(* IEC 61131-3 sources: plcassist-cli/packages/volt-lsp-iec/test-corpus/awa-palletizer/Device/Plc Logic/Application/Library Manager/VisuDialogs, 50 files *)

(* ---- DIALOG_CONSTANTS.gvl ---- *)
VAR_GLOBAL
	USERNAME_LABEL_DEFAULT : STRING := 'User';
	PASSWORD_LABEL_DEFAULT : STRING := 'Password';
	LOGIN_DIALOG_NAME : STRING := 'VisuDialogs.Login';
	PASSWORD_CHAR : STRING(1) := '*';
	CHAR_ASTERISK : BYTE := 42;
	CHAR_POINT : BYTE := 46;
	CHAR_SLASH : BYTE := 47;
	CHAR_BACKSLASH : BYTE := 92;
	ERR_DIR_NOT_FOUND : DWORD := 4000;
	ITFID_IGENERALCOMMAND : DWORD := 2;
	VISUDIALOGS_VERSION_ATLEAST_3_5_5 : INT := 0;
END_VAR

(* ---- DIALOG_VARIABLES.gvl ---- *)
VAR_GLOBAL
	G_FILELISTPROVIDER : Visu_FbFileListProvider;
	G_VISUDIALOGSCOMMANDS : Visu_DialogCommands;
END_VAR

(* ---- DIALOG_VARIABLES_EXP.gvl ---- *)
VAR_GLOBAL
	G_XEXP : BOOL;
END_VAR

(* ---- GVL_SORTEDFILELIST.gvl ---- *)
VAR_GLOBAL
	FILEELEMENTFACTORY : SortedDirectoryFileElementFactory;
	SORTEDLISTFACTORY : COL.SortedListFactory;
END_VAR

(* ---- IDIRECTORYFILEELEMENT.itf ---- *)
INTERFACE IDIRECTORYFILEELEMENT
END_INTERFACE

(* ---- IFILELISTPROVIDER.itf ---- *)
INTERFACE IFILELISTPROVIDER
END_INTERFACE

METHOD INITIALIZE : BOOL
VAR_INPUT
	STDIRECTORY : STRING(255);
	STFILTER : STRING;
	STFILEIN : STRING;
	STTITLE : STRING;
	IROWCOUNT : INT;
	BBROWSEDIRECTORY : BOOL;
	BTOUCH : BOOL;
END_VAR
END_METHOD

METHOD NEXT : BOOL
END_METHOD

METHOD PREVIOUS : BOOL
END_METHOD

(* ---- DIALOGCHECKINIT.fun ---- *)
FUNCTION DIALOGCHECKINIT : BOOL
VAR_IN_OUT
	STVALUE : STRING;
	STOUTPUT : STRING;
	BINIT : BOOL;
END_VAR
END_FUNCTION

(* ---- DIALOGCHECKINITFOREXPONENTIAL.fun ---- *)
FUNCTION DIALOGCHECKINITFOREXPONENTIAL : BOOL
VAR_INPUT
	STVALUE : STRING;
END_VAR
VAR_IN_OUT
	BINIT : BOOL;
END_VAR
END_FUNCTION

(* ---- DIALOGCHECKINITFOREXPONENTIALW.fun ---- *)
FUNCTION DIALOGCHECKINITFOREXPONENTIALW : BOOL
VAR_INPUT
	WSTVALUE : WSTRING;
END_VAR
VAR_IN_OUT
	BINIT : BOOL;
END_VAR
END_FUNCTION

(* ---- DIALOGCHECKINITW.fun ---- *)
FUNCTION DIALOGCHECKINITW : BOOL
VAR_IN_OUT
	WSTVALUE : WSTRING;
	WSTOUTPUT : WSTRING;
	BINIT : BOOL;
END_VAR
END_FUNCTION

(* ---- VISUDLG_CHECKEDAPPEND.fun ---- *)
FUNCTION VISUDLG_CHECKEDAPPEND : BOOL
VAR_INPUT
	BPASSWORD : BOOL;
	CTOAPPEND : STRING(1);
END_VAR
VAR_IN_OUT
	STOUTPUTVALUE : STRING;
	STVARIABLEVALUE : STRING;
	BINIT : BOOL;
END_VAR
END_FUNCTION

(* ---- VISUDLG_CHECKEDAPPENDEXP.fun ---- *)
FUNCTION VISUDLG_CHECKEDAPPENDEXP : BOOL
VAR_INPUT
	BPASSWORD : BOOL;
END_VAR
VAR_IN_OUT
	STOUTPUTVALUE : STRING;
	STVARIABLEVALUE : STRING;
	BINIT : BOOL;
END_VAR
END_FUNCTION

(* ---- VISUDLG_CHECKEDAPPENDW.fun ---- *)
FUNCTION VISUDLG_CHECKEDAPPENDW : BOOL
VAR_INPUT
	BPASSWORD : BOOL;
	CTOAPPEND : WSTRING(1);
END_VAR
VAR_IN_OUT
	WSTOUTPUTVALUE : WSTRING;
	WSTVARIABLEVALUE : WSTRING;
	BINIT : BOOL;
END_VAR
END_FUNCTION

(* ---- VISUDLG_CHECKEDBACK.fun ---- *)
FUNCTION VISUDLG_CHECKEDBACK : BOOL
VAR_IN_OUT
	STOUTPUTVALUE : STRING;
	STVARIABLEVALUE : STRING;
	BINIT : BOOL;
END_VAR
END_FUNCTION

(* ---- VISUDLG_CHECKEDBACKW.fun ---- *)
FUNCTION VISUDLG_CHECKEDBACKW : BOOL
VAR_IN_OUT
	WSTOUTPUTVALUE : WSTRING;
	WSTVARIABLEVALUE : WSTRING;
	BINIT : BOOL;
END_VAR
END_FUNCTION

(* ---- VISUDLG_CHECKEDCHANGENUMBERFORMAT.fun ---- *)
FUNCTION VISUDLG_CHECKEDCHANGENUMBERFORMAT : BOOL
VAR_INPUT
	BPASSWORD : BOOL;
	STCLICKEDRADIO : STRING;
END_VAR
VAR_IN_OUT
	STOUTPUTVALUE : STRING;
	STVARIABLEVALUE : STRING;
	STMIN : STRING;
	STMAX : STRING;
	IFORMATVALUE : INT;
END_VAR
END_FUNCTION

(* ---- VISUDLG_CHECKEDCHANGESIGN.fun ---- *)
FUNCTION VISUDLG_CHECKEDCHANGESIGN : BOOL
VAR_INPUT
	BPASSWORD : BOOL;
END_VAR
VAR_IN_OUT
	STOUTPUTVALUE : STRING;
	STVARIABLEVALUE : STRING;
	BINIT : BOOL;
END_VAR
END_FUNCTION

(* ---- VISUDLG_CHECKEDCHANGESIGNEXTENDED.fun ---- *)
FUNCTION VISUDLG_CHECKEDCHANGESIGNEXTENDED : BOOL
VAR_INPUT
	BPASSWORD : BOOL;
	IFORMATVALUE : INT;
END_VAR
VAR_IN_OUT
	STOUTPUTVALUE : STRING;
	STVARIABLEVALUE : STRING;
	BINIT : BOOL;
END_VAR
END_FUNCTION

(* ---- VISUDLG_CHECKEDCLEAR.fun ---- *)
FUNCTION VISUDLG_CHECKEDCLEAR : BOOL
VAR_IN_OUT
	STOUTPUTVALUE : STRING;
	STVARIABLEVALUE : STRING;
	FLAGS : DWORD;
END_VAR
END_FUNCTION

(* ---- VISUDLG_CHECKEDEXPFLOATFORMATSWITCH.fun ---- *)
FUNCTION VISUDLG_CHECKEDEXPFLOATFORMATSWITCH : BOOL
VAR_INPUT
	BPASSWORD : BOOL;
END_VAR
VAR_IN_OUT
	STOUTPUTVALUE : STRING;
	STVARIABLEVALUE : STRING;
END_VAR
END_FUNCTION

(* ---- VISUDLG_GETPASSWORDSTRING.fun ---- *)
FUNCTION VISUDLG_GETPASSWORDSTRING : STRING
VAR_INPUT
	STORG : STRING;
END_VAR
END_FUNCTION

(* ---- VISUDLG_PROCESSCHANGENUMBERFORMAT.fun ---- *)
FUNCTION VISUDLG_PROCESSCHANGENUMBERFORMAT : BOOL
VAR_INPUT
	BPASSWORD : BOOL;
	STCLICKEDRADIO : STRING;
END_VAR
VAR_IN_OUT
	STOUTPUTVALUE : STRING;
	STVARIABLEVALUE : STRING;
	STMIN : STRING;
	STMAX : STRING;
	IFORMATVALUE : INT;
	ICARETPOSITION : INT;
	ISELECTIONSTART : INT;
	ISELECTIONEND : INT;
END_VAR
END_FUNCTION

(* ---- VISUDLG_PROCESSCHANGESIGN.fun ---- *)
FUNCTION VISUDLG_PROCESSCHANGESIGN : BOOL
VAR_INPUT
	BPASSWORD : BOOL;
END_VAR
VAR_IN_OUT
	STOUTPUTVALUE : STRING;
	STVARIABLEVALUE : STRING;
	ICARETPOSITION : INT;
	ISELECTIONSTART : INT;
	ISELECTIONEND : INT;
END_VAR
END_FUNCTION

(* ---- VISUDLG_PROCESSCHANGESIGNEXTENDED.fun ---- *)
FUNCTION VISUDLG_PROCESSCHANGESIGNEXTENDED : BOOL
VAR_INPUT
	BPASSWORD : BOOL;
	IFORMATVALUE : INT;
END_VAR
VAR_IN_OUT
	STOUTPUTVALUE : STRING;
	STVARIABLEVALUE : STRING;
	ICARETPOSITION : INT;
	ISELECTIONSTART : INT;
	ISELECTIONEND : INT;
	BINIT : BOOL;
END_VAR
END_FUNCTION

(* ---- VISUDLG_PROCESSCLEAR.fun ---- *)
FUNCTION VISUDLG_PROCESSCLEAR : BOOL
VAR_IN_OUT
	STOUTPUTVALUE : STRING;
	STVARIABLEVALUE : STRING;
	FLAGS : DWORD;
	ICARETPOSITION : INT;
	ISELECTIONSTART : INT;
	ISELECTIONEND : INT;
END_VAR
END_FUNCTION

(* ---- VISUDLG_PROCESSEXP.fun ---- *)
FUNCTION VISUDLG_PROCESSEXP : BOOL
VAR_INPUT
	BPASSWORD : BOOL;
END_VAR
VAR_IN_OUT
	STOUTPUTVALUE : STRING;
	STVARIABLEVALUE : STRING;
	ICARETPOSITION : INT;
	ISELECTIONSTART : INT;
	ISELECTIONEND : INT;
	BINIT : BOOL;
END_VAR
END_FUNCTION

(* ---- VISUDLG_PROCESSEXPFLOATFORMATSWITCH.fun ---- *)
FUNCTION VISUDLG_PROCESSEXPFLOATFORMATSWITCH : BOOL
VAR_INPUT
	BPASSWORD : BOOL;
END_VAR
VAR_IN_OUT
	STOUTPUTVALUE : STRING;
	STVARIABLEVALUE : STRING;
	ICARETPOSITION : INT;
	ISELECTIONSTART : INT;
	ISELECTIONEND : INT;
	BINIT : BOOL;
END_VAR
END_FUNCTION

(* ---- VISUDLG_SETERRORCOLOR.fun ---- *)
FUNCTION VISUDLG_SETERRORCOLOR : DWORD
VAR_INPUT
	BERROR : BOOL;
END_VAR
END_FUNCTION

(* ---- VISUDLG_UTF8PASSWORDCARETPOSITION.fun ---- *)
FUNCTION VISUDLG_UTF8PASSWORDCARETPOSITION : INT
VAR_INPUT
	IRUNELEN : INT;
	STVARIABLE : STRING;
END_VAR
END_FUNCTION

(* ---- VISUDLG_UTF8RUNELEN.fun ---- *)
FUNCTION VISUDLG_UTF8RUNELEN : INT
VAR_INPUT
	STVARIABLEVALUE : STRING;
	IINDEX : INT;
END_VAR
END_FUNCTION

(* ---- VISUDLGUTIL_CLOSENUMPADEXTENDED.fun ---- *)
FUNCTION VISUDLGUTIL_CLOSENUMPADEXTENDED : BOOL
VAR_INPUT
	FLAGS : DWORD;
END_VAR
VAR_IN_OUT
	STOUTPUTVALUE : STRING;
	STVARIABLEVALUE : STRING;
	STMIN : STRING;
	STMAX : STRING;
	IFORMATVALUE : INT;
	BINITFORMATVALUE : BOOL;
END_VAR
END_FUNCTION

(* ---- VISUDLGUTIL_CLOSENUMPADEXTENDED2.fun ---- *)
FUNCTION VISUDLGUTIL_CLOSENUMPADEXTENDED2 : BOOL
VAR_INPUT
	FLAGS : DWORD;
END_VAR
VAR_IN_OUT
	STOUTPUTVALUE : STRING;
	STVARIABLEVALUE : STRING;
	STMIN : STRING;
	STMAX : STRING;
	IFORMATVALUE : INT;
	BINITFORMATVALUE : BOOL;
	ICARETPOSITION : INT;
	ISELECTIONSTART : INT;
	ISELECTIONEND : INT;
END_VAR
END_FUNCTION

(* ---- VISUDLGUTIL_FORMATEXPTOG.fun ---- *)
FUNCTION VISUDLGUTIL_FORMATEXPTOG : STRING
VAR_INPUT
	STVALUE : STRING;
END_VAR
END_FUNCTION

(* ---- VISUDLGUTIL_FORMATVALUETODEC.fun ---- *)
FUNCTION VISUDLGUTIL_FORMATVALUETODEC : STRING
VAR_INPUT
	STVARIABLEVALUE : STRING;
END_VAR
END_FUNCTION

(* ---- VISUDLGUTIL_FORMATVALUETOHEX.fun ---- *)
FUNCTION VISUDLGUTIL_FORMATVALUETOHEX : STRING
VAR_INPUT
	STVARIABLEVALUE : STRING;
END_VAR
END_FUNCTION

(* ---- VISUDLGUTIL_INITVALUEFROMFLAGS.fun ---- *)
FUNCTION VISUDLGUTIL_INITVALUEFROMFLAGS : INT
VAR_INPUT
	FLAGS : DWORD;
END_VAR
VAR_IN_OUT
	BINITFORMATVALUE : BOOL;
	IFORMATVALUE : INT;
END_VAR
END_FUNCTION

(* ---- VISUDLGUTIL_ISDIALOGOPEN.fun ---- *)
FUNCTION VISUDLGUTIL_ISDIALOGOPEN : BOOL
VAR_INPUT
	LOGINDIALOG : VisuElems.VisuElemBase.IVisualisationDialog;
	PVISUCLIENT : POINTER TO VisuElems.VisuElemBase.VisuStructClientData;
	DLGMAN : VisuElems.VisuElemBase.IDialogManager;
END_VAR
END_FUNCTION

(* ---- VISUDLGUTIL_SETBINITFORMATVALUE.fun ---- *)
FUNCTION VISUDLGUTIL_SETBINITFORMATVALUE : BOOL
VAR_INPUT
	STNEWVALUE : STRING;
END_VAR
VAR_IN_OUT
	BINITFORMATVALUE : BOOL;
END_VAR
END_FUNCTION

(* ---- VISUDLGUTIL_UPDATEOUTPUTVALUE.fun ---- *)
FUNCTION VISUDLGUTIL_UPDATEOUTPUTVALUE : BOOL
VAR_INPUT
	BPASSWORD : BOOL;
END_VAR
VAR_IN_OUT
	STOUTPUTVALUE : STRING;
	STVARIABLEVALUE : STRING;
END_VAR
END_FUNCTION

(* ---- GLOBALTEXTLIST.fb ---- *)
FUNCTION_BLOCK GLOBALTEXTLIST
VAR
	M_TEXTLISTFILE : STRING(255);
	_STNAMESPACE : STRING;
END_VAR
END_FUNCTION_BLOCK

(* ---- IMAGEPOOLDIALOGS.fb ---- *)
FUNCTION_BLOCK IMAGEPOOLDIALOGS
VAR
	M_STNAMESPACE : STRING(80);
	M_STHELPVARID : STRING;
	M_STHELPVARPATH : STRING(255);
	M_STHELP : STRING;
	M_REGISTERIMAGES : BOOL := TRUE;
END_VAR
END_FUNCTION_BLOCK

METHOD FB_INIT : BOOL
VAR_INPUT
	BINITRETAINS : BOOL;
	BINCOPYCODE : BOOL;
END_VAR
END_METHOD

METHOD FB_REINIT : BOOL
END_METHOD

METHOD FB_EXIT : BOOL
VAR_INPUT
	BINCOPYCODE : BOOL;
END_VAR
END_METHOD

(* ---- MINMAXLABELS.fb ---- *)
FUNCTION_BLOCK MINMAXLABELS
VAR
	M_TEXTLISTFILE : STRING(255);
	_STNAMESPACE : STRING;
END_VAR
END_FUNCTION_BLOCK

(* ---- SORTEDDIRECTORYFILEELEMENT.fb ---- *)
FUNCTION_BLOCK SORTEDDIRECTORYFILEELEMENT EXTENDS InstanceBase
VAR
	STFILENAME : STRING;
	DIRINFO : DirInfo;
	DIRECTORYINFO : POINTER TO DirInfo;
	FILENAME : POINTER TO STRING;
END_VAR
END_FUNCTION_BLOCK

METHOD DISPOSE : BOOL
END_METHOD

METHOD PRVINSTINIT : FBF.Error
VAR_INPUT
	ITFDATA : FBF.IData;
END_VAR
END_METHOD

METHOD ELEMENTCOMPARETO : INT
VAR_INPUT
	ITFELEMENT : COL.IElement;
END_VAR
END_METHOD

METHOD ELEMENTEQUALS : BOOL
VAR_INPUT
	ITFELEMENT : COL.IElement;
END_VAR
END_METHOD

METHOD ELEMENTHASHCODE : LINT
END_METHOD

(* ---- SORTEDDIRECTORYFILEELEMENTDATA.fb ---- *)
FUNCTION_BLOCK SORTEDDIRECTORYFILEELEMENTDATA EXTENDS InstanceData
VAR_INPUT
	STFILENAME : STRING;
	DIRINFO : DirInfo;
END_VAR
END_FUNCTION_BLOCK

(* ---- SORTEDDIRECTORYFILEELEMENTFACTORY.fb ---- *)
FUNCTION_BLOCK SORTEDDIRECTORYFILEELEMENTFACTORY EXTENDS FactoryBase
VAR
	PRVINSTCOUNT : CAA.COUNT;
	PRVINSTPOOLEXTENDSFACTOR : USINT;
	PRVINSTSIZE : CAA.SIZE;
END_VAR
END_FUNCTION_BLOCK

METHOD CREATE : IDirectoryFileElement
VAR_INPUT
	STFILENAME : STRING;
	DIRINFO : DirInfo;
END_VAR
VAR_OUTPUT
	EERROR : FBF.ERROR;
END_VAR
END_METHOD

(* ---- VISU_DIALOGCOMMANDS.fb ---- *)
FUNCTION_BLOCK VISU_DIALOGCOMMANDS
VAR
	_CMDOPENFILEDIALOG : Visu_FbOpenFileDialog;
END_VAR
END_FUNCTION_BLOCK

METHOD FB_INIT
VAR_INPUT
	BINITRETAINS : BOOL;
	BINCOPYCODE : BOOL;
END_VAR
END_METHOD

METHOD REGISTERCOMMANDS : BOOL
VAR_INPUT
	COMMANDMANAGER : VisuElems.ICommandManager2;
END_VAR
END_METHOD

(* ---- VISU_FBDIALOGLOGINPROVIDER.fb ---- *)
FUNCTION_BLOCK VISU_FBDIALOGLOGINPROVIDER
VAR
	_STPASSWORD : STRING;
	_STUSERNAME : STRING;
	_CREDENTIALS : Visu_UserPasswordCredentials;
	_STTITLEPREFIX : STRING;
	_STCURRENTDATASOURCE : STRING;
	_STUSERLABELTEXT : STRING;
	_STPASSWORDLABELTEXT : STRING;
	_UXIPROVIDINGCREDENTIALSFOR : __UXINT;
	_UXINEXTREQUESTID : __UXINT;
	_RETRYWAITTIME : TIME;
	_UDIRETRYCOUNTER : UDINT;
	_UDIRETRIESPOSSIBLE : UDINT;
	_ITFICREDENTIALSPROVIDER : IDatasources.ICredentialsProvider := THIS^;
	_BDIALOGOPEN : BOOL;
	_BDIALOGRESULTAVAILABLE : BOOL;
	_BDIALOGACCEPTED : BOOL;
	_PCLIENTOPENEDDIALOGFOR : POINTER TO BYTE;
	DIALOGMAN : VisuElems.VisuElemBase.IDialogManager;
	LOGINDIALOG : VisuElems.VisuElemBase.IVisualisationDialog;
	PLOGININFO : POINTER TO Login_VISU_STRUCT;
	PVISUCLIENT : POINTER TO VisuElems.VisuElemBase.VisuStructClientData;
	RESULT : VisuElems.VisuElemBase.Visu_DialogResult;
	PASSWORD : STRING;
	PASSWORDLABELTEXT : STRING;
	RETRYWAITTIME : TIME;
	RETRYWAITTIME_MS : UDINT;
	TITLE : STRING;
	TITLEPREFIX : STRING;
	TRIALCOUNT : UDINT;
	USERLABELTEXT : STRING;
END_VAR
END_FUNCTION_BLOCK

METHOD GETCREDENTIALS : IDatasources.SysTypes.RTS_IEC_RESULT
VAR_INPUT
	UXIREQUESTID : __UXINT;
END_VAR
VAR_OUTPUT
	CREDENTIALS : IDatasources.ICredentials;
END_VAR
END_METHOD

METHOD ISGETCREDENTIALSFINISHED : IDatasources.SysTypes.RTS_IEC_RESULT
VAR_INPUT
	UXIREQUESTID : __UXINT;
END_VAR
END_METHOD

METHOD ISLOGINALREADOPEN : BOOL
VAR_INPUT
	LOGINDIALOG : VisuElems.VisuElemBase.IVisualisationDialog;
	PVISUCLIENT : POINTER TO VisuElems.VisuElemBase.VisuStructClientData;
	DLGMAN : VisuElems.VisuElemBase.IDialogManager;
END_VAR
END_METHOD

METHOD LOGINFAILED : UDINT
VAR_INPUT
	UXIREQUESTID : __UXINT;
END_VAR
VAR_OUTPUT
	TRETRYWAITTIME : TIME;
END_VAR
END_METHOD

METHOD LOGINSUCCEEDED
VAR_INPUT
	UXIREQUESTID : __UXINT;
END_VAR
END_METHOD

METHOD STARTGETCREDENTIALS : __UXINT
VAR_INPUT
	PSTDATASOURCE : POINTER TO STRING;
END_VAR
VAR_OUTPUT
	UDIERRORCODE : IDatasources.SysTypes.RTS_IEC_RESULT;
END_VAR
END_METHOD

METHOD PRVRESET : BOOL
END_METHOD

(* ---- VISU_FBFILELISTPROVIDER.fb ---- *)
FUNCTION_BLOCK VISU_FBFILELISTPROVIDER
VAR_INPUT
	STFILE : STRING;
END_VAR
VAR
	_STDIRECTORY : STRING(255);
	_STFILTER : STRING;
	_STFILTERDISPLAY : STRING;
	_STTITLE : STRING := 'Load file';
	_STOK : STRING(10) := 'Load';
	_BBROWSEDIRECTORY : BOOL := FALSE;
	_BCHANGESELECTION : BOOL := FALSE;
	_STLFILES : ARRAY [0..MAX_FILE_NAMES] OF STRING;
	_STLIMAGES : ARRAY [0..MAX_FILE_NAMES] OF STRING(3);
	_STDIRECTORYFILTER : STRING(255);
	_STNEWFOLDER : STRING(255);
	_PSTNEWFOLDER : POINTER TO STRING;
	_IFILES : INT;
	_IINDEX : INT;
	_IINDEXSLIDER : INT;
	_IPREVINDEXSLIDER : INT;
	_IROWCOUNT : INT;
	_ISELECTIONINDEX : INT := -1;
	_IPREVSELECTIONINDEX : INT := -1;
	_IPREVPREVSELECTIONINDEX : INT;
	_DWLASTERROR : DWORD;
	_BDELETE : BOOL := FALSE;
	_BDIRUP : BOOL := FALSE;
	_BTOUCH : BOOL := TRUE;
	_BDIRSELECTED : BOOL;
	ILEN : INT;
	IPOS : INT;
	IARRAYINDEX : INT;
	BROOTDIRISSLASH : BOOL := FALSE;
	MAX_FILE_NAMES : INT := 12;
	COUNT : INT;
END_VAR
END_FUNCTION_BLOCK

METHOD DUMMY : INT
END_METHOD

METHOD GETSELECTEDDIRECTORY : STRING
END_METHOD

METHOD GETSELECTEDFILENAME : STRING
END_METHOD

METHOD INITIALIZE : BOOL
VAR_INPUT
	STDIRECTORY : STRING(255);
	STFILTER : STRING;
	STFILEIN : STRING;
	STTITLE : STRING;
	IROWCOUNT : INT;
	BBROWSEDIRECTORY : BOOL;
	BTOUCH : BOOL;
END_VAR
END_METHOD

METHOD NEXT : BOOL
END_METHOD

METHOD PREVIOUS : BOOL
END_METHOD

METHOD PRVADD : BOOL
VAR_INPUT
	STFILE : STRING;
	PIFILEINDEX : POINTER TO INT;
	PIARRAYINDEX : POINTER TO INT;
	PDIRINFO : POINTER TO DirInfo;
	BONLYFOLDER : BOOL;
END_VAR
END_METHOD

METHOD PRVADDFILEFILTERED : BOOL
VAR_IN_OUT
	ITFDIRECTORYFILEELEM : IDirectoryFileElement;
	IFILEINDEX : INT;
	IARRAYINDEX : INT;
	XNOFILTER : BOOL;
	PSTFILTERHELP : POINTER TO STRING;
	ILENFILTER : INT;
END_VAR
END_METHOD

METHOD PRVCLEAR : BOOL
END_METHOD

METHOD PRVCOLLECTFILES : BOOL
VAR_IN_OUT
	SORTEDLIST : COL.ISortedList2;
END_VAR
END_METHOD

METHOD PRVRESETINDEX : BOOL
END_METHOD

METHOD PRVSEARCH : BOOL
END_METHOD

(* ---- VISU_FBOPENFILEDIALOG.fb ---- *)
FUNCTION_BLOCK VISU_FBOPENFILEDIALOG
VAR
	_ITFGENERALCOMMAND : VisuElems.IGeneralCommand2 := THIS^;
	_PDLGPARAMS : POINTER TO VisuElems.Visu_StructVisuFileDialogParams;
	ROW_COUNT : INT := 6;
END_VAR
END_FUNCTION_BLOCK

METHOD EXECUTE : __XWORD
VAR_INPUT
	DWPARAM1 : __XWORD;
	DWPARAM2 : __XWORD;
END_VAR
END_METHOD

METHOD GETINTERFACE : POINTER TO BYTE
VAR_INPUT
	DWITFID : DWORD;
END_VAR
END_METHOD

(* ---- VISU_USERPASSWORDCREDENTIALS.fb ---- *)
FUNCTION_BLOCK VISU_USERPASSWORDCREDENTIALS
VAR_INPUT
	STPASSWORD : STRING;
	STUSERNAME : STRING;
END_VAR
VAR
	PASSWORD : STRING;
	USERNAME : STRING;
END_VAR
END_FUNCTION_BLOCK
